Universal Robots URScript: T011_zai-org_GLM-4.7-FP8_baseline_rep3.urscript

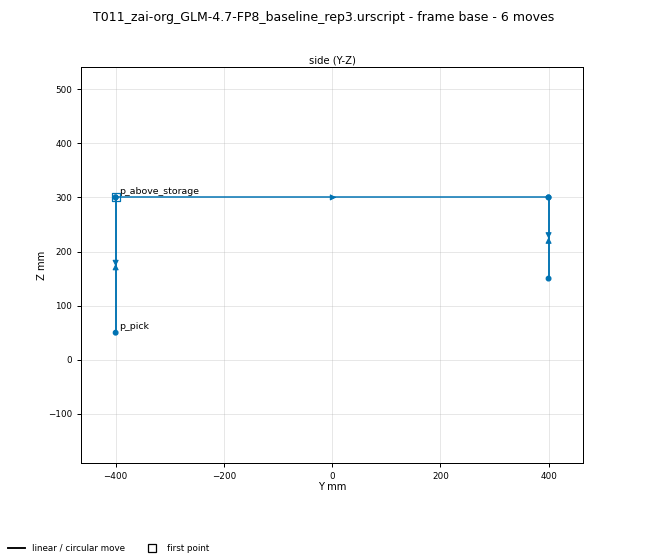
[picture p0: tool path of T011_zai-org_GLM-4.7-FP8_baseline_rep3.urscript in frame base, 6 of 8 moves have a stored position in this frame; points joined in program order, loops and branches not executed]
# Program: Dual-zone pick-place — hybrid mode (T011)
# Robot: UR5e
# Payload: 1.2 kg

# Configuration
set_payload(1.2, [0.0, 0.0, 0.0])
set_tcp(p[0.0, 0.0, 0.0, 0.0, 0.0, 0.0])

# Waypoint Definitions
q_home = [0.0, -1.57, 0.0, -1.57, 0.0, 0.0]

# Storage Zone (Fenced)
p_above_storage = p[0.4, -0.4, 0.3, 3.14, 0.0, 0.0]
p_pick = p[0.4, -0.4, 0.05, 3.14, 0.0, 0.0]

# Handoff Zone (Collaborative)
p_above_handoff = p[0.4, 0.4, 0.3, 3.14, 0.0, 0.0]
p_handoff = p[0.4, 0.4, 0.15, 3.14, 0.0, 0.0]

# --- Motion Sequence ---

# 1. Move Joint: Home, 250.0 mm/s
movej(q_home, a=1.2, v=0.25)

# 2. Move Linear: Above storage bin, 280.0 mm/s
# Entering Safety Zone: Confinement
movel(p_above_storage, a=1.0, v=0.28)

# 3. Move Linear: Descend to pick, 120.0 mm/s
movel(p_pick, a=0.5, v=0.12)

# Action: Gripper Close
set_tool_digital_out(0, True)
sleep(0.5)

# 4. Move Linear: Lift from bin, 200.0 mm/s
movel(p_above_storage, a=0.8, v=0.20)

# 5. Move Linear: Transit to handoff zone, 250.0 mm/s
# Transitioning to Collaborative Zone
# Entering Safety Zone: Exclusion (Operator area)
movel(p_above_handoff, a=1.0, v=0.25)

# 6. Move Linear: Descend to handoff, 100.0 mm/s (Slower for safety)
movel(p_handoff, a=0.5, v=0.10)

# Action: Gripper Open
set_tool_digital_out(0, False)
sleep(0.5)

# 7. Move Linear: Lift from handoff, 200.0 mm/s
movel(p_above_handoff, a=0.8, v=0.20)

# 8. Move Joint: Return Home, 250.0 mm/s
movej(q_home, a=1.2, v=0.25)

# End of Program
